// TIA Portal V19 export
TYPE "AnaMon.Feature"
   STRUCT
      Startup : Bool := TRUE;
   END_STRUCT;
END_TYPE
